FUNCTION_BLOCK fb_Dev_AnalogSensor_ELM_10x EXTENDS fb_Dev_AnalogSensor
VAR_INPUT
	inpRawIOChannelArray			: ARRAY [1..10] OF DINT;
END_VAR
VAR_OUTPUT
	stsSensorRawSignalArray	: ARRAY [1..10] OF LREAL;
	stsEngValueArray		: ARRAY [1..10] OF LREAL;
	stsEngValueRMS			: LREAL;
END_VAR
VAR
	_sensorRawSignalArray			: ARRAY [1..10] OF LREAL;
	_engValueArray					: ARRAY [1..10] OF LREAL;
	_engValueRMS					: LREAL;
END_VAR

// This FB is intended for a ELM IO card set to 10x overscan with a 1ms CPU cycletime

DeviceLogic();

scaleInput();

FaultHandler();

setHMI();

stsSensorRawSignalArray		:= _sensorRawSignalArray;
stsEngValueArray			:= _engValueArray;

stsSensorRawSignal 			:= _sensorRawSignal;
stsEngValue					:= _engValue;

METHOD scaleInput : BOOL
VAR
	i : INT;
	tempRaw : LREAL := 0.0;
	tempEng : LREAL := 0.0;
	tempEngSqSum 	: LREAL := 0.0;
END_VAR
FOR i := 1 TO 10 DO
	_sensorRawSignalArray[i]	:= F_AnalogToEngUnit(inpRawIOChannelArray[i], cfgChannelMinInt, cfgChannelMaxInt, cfgSensorMin, cfgSensorMax);
	_engValueArray[i]			:= (F_AnalogToEngUnit(_sensorRawSignalArray[i], cfgSensorMin, cfgSensorMax, cfgEngUnitMin, cfgEngUnitMax) * _CalGain) + _CalOffset;
	tempRaw := tempRaw + _sensorRawSignalArray[i];
	tempEng := tempEng + _engValueArray[i];
	tempEngSqSum := tempEngSqSum + _engValueArray[i] * _engValueArray[i];
END_FOR

_sensorRawSignal	:= tempRaw / 10;
_engValue			:= tempEng / 10;
_engValueRMS		:= SQRT(tempEngSqSum / 10);
END_METHOD

END_FUNCTION_BLOCK

(* stored: Version 1.1.0.1
   POU fb_Dev_AnalogSensor_ELM_10x: Id {02f7c873-b950-4330-818a-26fa0d414421}, SpecialFunc None
   Method scaleInput: Id {c81df925-397f-4824-b11a-b5153ad9d3c9} *)
